FUNCTION_BLOCK E_SELECT_5 (* Extracted Composite Function Block Type *)
  (* Standard: 61499-2 *)
  (* Version 10/22/2026, macie *)
  PACKAGE Main;
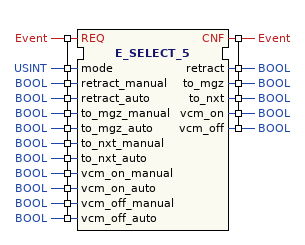
  EVENT_INPUT
    REQ WITH mode, retract_manual, retract_auto, to_mgz_manual, to_mgz_auto, to_nxt_manual, to_nxt_auto, vcm_on_manual, vcm_on_auto, vcm_off_manual, vcm_off_auto; (* Normal Execution Request *)
  END_EVENT
  EVENT_OUTPUT
    CNF WITH retract, to_mgz, to_nxt, vcm_on, vcm_off; (* Execution Confirmation *)
  END_EVENT
  VAR_INPUT
    mode : USINT; (* Selector *)
    retract_manual : BOOL; (* Argument *)
    retract_auto : BOOL; (* Argument *)
    to_mgz_manual : BOOL; (* Argument *)
    to_mgz_auto : BOOL; (* Argument *)
    to_nxt_manual : BOOL; (* Argument *)
    to_nxt_auto : BOOL; (* Argument *)
    vcm_on_manual : BOOL; (* Argument *)
    vcm_on_auto : BOOL; (* Argument *)
    vcm_off_manual : BOOL; (* Argument *)
    vcm_off_auto : BOOL; (* Argument *)
  END_VAR
  VAR_OUTPUT
    retract : BOOL; (* Result: IN1 or IN2 or ... according to the SELECT input (SELECT = 0 selects IN1) *)
    to_mgz : BOOL; (* Result: IN1 or IN2 or ... according to the SELECT input (SELECT = 0 selects IN1) *)
    to_nxt : BOOL; (* Result: IN1 or IN2 or ... according to the SELECT input (SELECT = 0 selects IN1) *)
    vcm_on : BOOL; (* Result: IN1 or IN2 or ... according to the SELECT input (SELECT = 0 selects IN1) *)
    vcm_off : BOOL; (* Result: IN1 or IN2 or ... according to the SELECT input (SELECT = 0 selects IN1) *)
  END_VAR
  FBS
    SELECT_RETRACT : SELECT_783952938E11160B; {SET_ATTRIBUTE(Configuration.GenericFBType.InterfaceParams, Runtime.Standard#CNT:=2;IN${CNT$}:BOOL)}
    SELECT_TO_MGZ : SELECT_783952938E11160B; {SET_ATTRIBUTE(Configuration.GenericFBType.InterfaceParams, Runtime.Standard#CNT:=2;IN${CNT$}:BOOL)}
    SELECT_TO_NXT : SELECT_783952938E11160B; {SET_ATTRIBUTE(Configuration.GenericFBType.InterfaceParams, Runtime.Standard#CNT:=2;IN${CNT$}:BOOL)}
    SELECT_VCM_ON : SELECT_783952938E11160B; {SET_ATTRIBUTE(Configuration.GenericFBType.InterfaceParams, Runtime.Standard#CNT:=2;IN${CNT$}:BOOL)}
    SELECT_VCM_OFF : SELECT_783952938E11160B; {SET_ATTRIBUTE(Configuration.GenericFBType.InterfaceParams, Runtime.Standard#CNT:=2;IN${CNT$}:BOOL)}
  END_FBS
  EVENT_CONNECTIONS
    SELECT_RETRACT.CNF TO CNF;
    REQ TO SELECT_RETRACT.REQ;
    REQ TO SELECT_TO_MGZ.REQ;
    REQ TO SELECT_TO_NXT.REQ;
    REQ TO SELECT_VCM_ON.REQ;
    REQ TO SELECT_VCM_OFF.REQ;
  END_CONNECTIONS
  DATA_CONNECTIONS
    mode TO SELECT_RETRACT.SELECT;
    retract_manual TO SELECT_RETRACT.IN1;
    retract_auto TO SELECT_RETRACT.IN2;
    SELECT_RETRACT.OUT TO retract;
    to_mgz_manual TO SELECT_TO_MGZ.IN1;
    to_mgz_auto TO SELECT_TO_MGZ.IN2;
    SELECT_TO_MGZ.OUT TO to_mgz;
    to_nxt_manual TO SELECT_TO_NXT.IN1;
    to_nxt_auto TO SELECT_TO_NXT.IN2;
    SELECT_TO_NXT.OUT TO to_nxt;
    vcm_on_manual TO SELECT_VCM_ON.IN1;
    vcm_on_auto TO SELECT_VCM_ON.IN2;
    SELECT_VCM_ON.OUT TO vcm_on;
    vcm_off_manual TO SELECT_VCM_OFF.IN1;
    vcm_off_auto TO SELECT_VCM_OFF.IN2;
    SELECT_VCM_OFF.OUT TO vcm_off;
    mode TO SELECT_VCM_OFF.SELECT;
    mode TO SELECT_TO_MGZ.SELECT;
    mode TO SELECT_TO_NXT.SELECT;
    mode TO SELECT_VCM_ON.SELECT;
  END_CONNECTIONS
END_FUNCTION_BLOCK
